DATA_BLOCK "naut_SfcStepT_DB"
{ S7_Optimized_Access := 'TRUE' }
VERSION : 0.1
"naut_SfcStepT"

BEGIN

END_DATA_BLOCK
